// TIA Portal V20 export
TYPE "AZ_PrmRW_PLC2Drv"
   STRUCT
      ReadParameterID : Word;
      WriteRequest : Struct
         Reserved_32 : Byte;
         "WR-REQ" : Bool;
         Reserved_33_bit1 : Bool;
         Reserved_33_bit2 : Bool;
         Reserved_33_bit3 : Bool;
         Reserved_33_bit4 : Bool;
         Reserved_33_bit5 : Bool;
         Reserved_33_bit6 : Bool;
         Reserved_33_bit7 : Bool;
      END_STRUCT;
      WriteParameterID : Word;
      WriteData : DInt;
   END_STRUCT;
END_TYPE
